RoboDK station: FlowControlTest_oficial.rdk

Station FlowControlTest (saved by RoboDK 5.6.5). Poses are relative to the parent item; angles as X-Y-Z fixed-axis rotations.
Station parameters (name, value as stored): CNC1_DoorClosed , 1, CNC1_DoorOpened , 0, CNC1_CloseDoor , 1, CNC1_CloseDoor, 1
  - program SetOpenDoor (1 instructions, listed below)
  - program SetCloseDoor (1 instructions, listed below)
  - program Program1 (8 instructions, listed below)
  - program CloseDoor (2 instructions, listed below)

--- program SetOpenDoor ---
  Set CNC1_CloseDoor=0

--- program SetCloseDoor ---
  Set CNC1_CloseDoor=1

--- program Program1 ---
  IF CNC1_CloseDoor == 1
  Call CloseDoor
  Set CNC1_DoorClosed =1
  Set CNC1_DoorOpened =0
  ELSE: END
  Print: DOOR ALREADY CLOSED!
  Stop
  END

--- program CloseDoor ---
  Print: CLOSING DOOR!
  Stop
